(****************************************************************************************************<br>
© Syntegon Group.<br>
All rights reserved, also regarding any disposal, exploitation, reproduction, editing, distribution,<br>
as well as in the event of applications for industrial property rights.<br>
*****************************************************************************************************<br>
DESCRIPTION:<br>
Parameter set of one XTS loop (ADR 0017): its pose, origin shift, track modules, zones and gripper fingers,<br>
written by the configurator, taken over when the application allows it. Typical cycle:<br>
  fb_FxxParam.m_Register(vio_Manifest := GVL_Config.stManifest, vi_udn_Id := fb_Fxx.m_Id());<br>
  fb_FxxParam.m_Cycle(vio_Default := FxxDefault, vio_Set := FxxSet, vi_b_ApplyAllowed := b_Stopped);<br>
  fb_Fxx.m_Configure(vi_lr_ToolOffset := 120, ...);<br>
  fb_FxxParam.m_PassOn(vio_Visu := fb_Fxx);<br>
The application's logic takes its track and zones from m_Active, not from its own constants.<br>
*****************************************************************************************************<br>
OUTPUT VALUES:<br>
vo_Config is the contract structure the gateway reads and writes at the path in the config manifest.<br>
*****************************************************************************************************<br>
VERSION         ¦ DATE       ¦ NAME      ¦ CHANGE<br>
Syn_Config 1.1.0 ¦ 2026-11-10 ¦ J.Willner ¦ New<br>
Syn_Config 2.0.0 ¦ 2026-11-11 ¦ J.Willner ¦ Gripper fingers with their offsets (ADR 0018)<br>
Syn_Config 2.3.0 ¦ 2026-11-14 ¦ J.Willner ¦ m_Cycle through m_HandleStaging; m_PassOn passes the pose on<br>
****************************************************************************************************)
FUNCTION_BLOCK _FB_ConfigXtsLoop EXTENDS _FB_ConfigComponent
VAR_OUTPUT
	vo_Config							: ST_ConfigXtsLoop;	// contract structure of the gateway
END_VAR

(****************************************************************************************************<br>
© Syntegon Group.<br>
All rights reserved, also regarding any disposal, exploitation, reproduction, editing, distribution,<br>
as well as in the event of applications for industrial property rights.<br>
*****************************************************************************************************<br>
DESCRIPTION:<br>
All effective values (track modules, zones, ...), for the application's own logic.<br>
****************************************************************************************************)
METHOD m_Active : ST_ConfigXtsLoopParam
m_Active := vo_Config.stActive;
END_METHOD

(****************************************************************************************************<br>
© Syntegon Group.<br>
All rights reserved, also regarding any disposal, exploitation, reproduction, editing, distribution,<br>
as well as in the event of applications for industrial property rights.<br>
*****************************************************************************************************<br>
DESCRIPTION:<br>
An XTS loop.<br>
****************************************************************************************************)
METHOD PROTECTED m_ComponentType : SynVisu.E_VisuComponentType
m_ComponentType := SynVisu.E_VisuComponentType.XTS_LOOP;
END_METHOD

(****************************************************************************************************<br>
© Syntegon Group.<br>
All rights reserved, also regarding any disposal, exploitation, reproduction, editing, distribution,<br>
as well as in the event of applications for industrial property rights.<br>
*****************************************************************************************************<br>
DESCRIPTION:<br>
Every cycle: handles a staged set or a reset (a set only while vi_b_ApplyAllowed), keeps the active set in<br>
vio_Set and gives the effective values in vo_Config.stActive: the active set while one is valid, else the<br>
program values vio_Default.<br>
*****************************************************************************************************<br>
OUTPUT VALUES:<br>
TRUE in the cycle a set was taken over or reset.<br>
****************************************************************************************************)
METHOD m_Cycle : BOOL
VAR_IN_OUT CONSTANT
	vio_Default							: ST_ConfigXtsLoopParam;	// the application's program values
END_VAR
VAR_IN_OUT
	vio_Set								: ST_ConfigXtsLoopSet;	// the application's VAR PERSISTENT active set
END_VAR
VAR_INPUT
	vi_b_ApplyAllowed					: BOOL;	// [-] a staged set may be taken over now, e.g. while the machine stands
END_VAR
VAR
	b_TempTakeOver						: BOOL;	// the staged set was taken over: copy it
END_VAR
m_Cycle := m_HandleStaging(vio_Staging := vo_Config.stStaging, vio_Status := vo_Config.stStatus, vio_b_Valid := vio_Set.bValid,
	vio_udn_Version := vio_Set.nVersion, vio_udn_LastVersion := vio_Set.nLastVersion, vi_b_ApplyAllowed := vi_b_ApplyAllowed,
	vo_b_TakeOver => b_TempTakeOver);
IF b_TempTakeOver THEN
	vio_Set.stParam := vo_Config.stStaged;
END_IF


(****************************************************************************************************
EFFECTIVE VALUES
****************************************************************************************************)
IF vio_Set.bValid THEN
	vo_Config.stActive := vio_Set.stParam;
ELSE
	vo_Config.stActive := vio_Default;
END_IF
END_METHOD

(****************************************************************************************************<br>
© Syntegon Group.<br>
All rights reserved, also regarding any disposal, exploitation, reproduction, editing, distribution,<br>
as well as in the event of applications for industrial property rights.<br>
*****************************************************************************************************<br>
DESCRIPTION:<br>
Why a staged set cannot be taken over; '' when it can: a track without modules, more modules, zones or fingers<br>
than the lists hold, a module without a length, a zone on no conveyor (id 0), or a finger without a diameter or<br>
height.<br>
****************************************************************************************************)
METHOD PROTECTED m_InvalidStaged : STRING(80)
m_InvalidStaged := m_InvalidModules(vio_aModules := vo_Config.stStaged.aModules, vi_un_Count := vo_Config.stStaged.nModuleCount);
IF m_InvalidStaged = '' THEN
	m_InvalidStaged := m_InvalidZones(vio_aZones := vo_Config.stStaged.aZones, vi_un_Count := vo_Config.stStaged.nZoneCount);
END_IF
IF m_InvalidStaged = '' THEN
	m_InvalidStaged := m_InvalidFingers(vio_aFingers := vo_Config.stStaged.aFingers, vi_un_Count := vo_Config.stStaged.nFingerCount);
END_IF
END_METHOD

(****************************************************************************************************<br>
© Syntegon Group.<br>
All rights reserved, also regarding any disposal, exploitation, reproduction, editing, distribution,<br>
as well as in the event of applications for industrial property rights.<br>
*****************************************************************************************************<br>
DESCRIPTION:<br>
Passes the effective pose, origin shift, track modules, zones and fingers on to the loop's Syn_Visu FB, so the<br>
visualisation shows what the machine uses; the tool offset and mover size (hardware) stay with the<br>
application's m_Configure call. Call it after m_Cycle, every cycle; Syn_Visu's config version only changes when<br>
a value does.<br>
****************************************************************************************************)
METHOD m_PassOn : BOOL
VAR_IN_OUT
	vio_Visu							: SynVisu._FB_VisuXtsLoop;	// the loop's Syn_Visu FB
END_VAR
m_PassOn := TRUE;
vio_Visu.m_SetPose(vi_Pose := vo_Config.stActive.stPose);
vio_Visu.m_SetOriginShift(vi_lr_X := vo_Config.stActive.stOriginShift.fX, vi_lr_Y := vo_Config.stActive.stOriginShift.fY,
	vi_lr_Z := vo_Config.stActive.stOriginShift.fZ);
m_PassOnModules(vio_Visu := vio_Visu, vio_aModules := vo_Config.stActive.aModules,
	vi_un_Count := vo_Config.stActive.nModuleCount, vi_un_VisuCount := vio_Visu.vo_Visu.stConfig.nModuleCount);
m_PassOnZones(vio_Visu := vio_Visu, vio_aZones := vo_Config.stActive.aZones, vi_un_Count := vo_Config.stActive.nZoneCount,
	vi_un_VisuCount := vio_Visu.vo_Visu.stConfig.nZoneCount);
m_PassOnFingers(vio_Visu := vio_Visu, vio_aFingers := vo_Config.stActive.aFingers,
	vi_un_Count := vo_Config.stActive.nFingerCount, vi_un_VisuCount := vio_Visu.vo_Visu.stConfig.nFingerCount);
END_METHOD

(****************************************************************************************************<br>
© Syntegon Group.<br>
All rights reserved, also regarding any disposal, exploitation, reproduction, editing, distribution,<br>
as well as in the event of applications for industrial property rights.<br>
*****************************************************************************************************<br>
DESCRIPTION:<br>
Effective pose of the start of module 1 (MCS), for the application's logic.<br>
****************************************************************************************************)
METHOD m_Pose : SynVisu.ST_VisuPose
m_Pose := vo_Config.stActive.stPose;
END_METHOD

END_FUNCTION_BLOCK

(* stored: Version 1.1.0.1
   POU _FB_ConfigXtsLoop: Id {0dc8dfc6-59a5-4dff-95a7-eb94b158a9f9}, SpecialFunc None
   Method m_Active: Id {1f24dc3b-afdd-46cf-b338-33bd7aa3e73e}
   Method m_ComponentType: Id {243d541e-cb5a-4823-8566-8fd186b7d04d}
   Method m_Cycle: Id {abf9ad5a-3af4-42e0-9821-0f5b09453a7e}
   Method m_InvalidStaged: Id {2b281ea4-5528-4ad1-9b1b-c40296c7e24f}
   Method m_PassOn: Id {22d4fb07-6885-4daa-9d98-da72bba0c32d}
   Method m_Pose: Id {eec44d82-e17a-42a6-b9be-483f3ceaf7fe} *)
